(* IEC 61131-3 sources: TSA-FMICS22/ahorn/test/lib_se/file, 7 files *)

(* ---- call_coverage_in_1_cycle_with_change_annotation.st ---- *)
PROGRAM P
VAR_INPUT
    a : INT;
END_VAR
VAR
    f : Fb;
END_VAR
VAR_OUTPUT
    b : BOOL;
END_VAR
    f(x:=a,z=>b);
END_PROGRAM

FUNCTION_BLOCK Fb
VAR_INPUT
    x : INT;
END_VAR
VAR
    y : INT;
END_VAR
VAR_OUTPUT
    z : BOOL;
END_VAR;
    IF x >= 32 THEN
        y := y + change(1, 3);
    ELSE
        y := y;
    END_IF;
    IF y >= 3 THEN
        z := TRUE;
        y := 0;
    ELSE
        z := FALSE;
    END_IF;
END_FUNCTION_BLOCK

(* ---- call_coverage_in_2_cycles.st ---- *)
PROGRAM P
VAR_INPUT
    a : INT;
END_VAR
VAR
    f : Fb;
END_VAR
VAR_OUTPUT
    b : BOOL;
END_VAR
    f(x:=a,z=>b);
END_PROGRAM

FUNCTION_BLOCK Fb
VAR_INPUT
    x : INT;
END_VAR
VAR
    y : INT;
END_VAR
VAR_OUTPUT
    z : BOOL;
END_VAR;
    IF x >= 32 THEN
        y := y + 2;
    ELSE
        y := y;
    END_IF;
    IF y >= 3 THEN
        z := TRUE;
        y := 0;
    ELSE
        z := FALSE;
    END_IF;
END_FUNCTION_BLOCK

(* ---- call_coverage_in_2_cycles_with_change_annotation.st ---- *)
PROGRAM P
VAR_INPUT
    a : INT;
END_VAR
VAR
    f : Fb;
END_VAR
VAR_OUTPUT
    b : BOOL;
END_VAR
    f(x:=a,z=>b);
END_PROGRAM

FUNCTION_BLOCK Fb
VAR_INPUT
    x : INT;
END_VAR
VAR
    y : INT;
END_VAR
VAR_OUTPUT
    z : BOOL;
END_VAR;
    IF x >= 32 THEN
        y := y + change(1, 2);
    ELSE
        y := y;
    END_IF;
    IF y >= 3 THEN
        z := TRUE;
        y := 0;
    ELSE
        z := FALSE;
    END_IF;
END_FUNCTION_BLOCK

(* ---- call_coverage_in_3_cycles.st ---- *)
PROGRAM P
VAR_INPUT
    a : INT;
END_VAR
VAR
    f : Fb;
END_VAR
VAR_OUTPUT
    b : BOOL;
END_VAR
    f(x:=a,z=>b);
END_PROGRAM

FUNCTION_BLOCK Fb
VAR_INPUT
    x : INT;
END_VAR
VAR
    y : INT;
END_VAR
VAR_OUTPUT
    z : BOOL;
END_VAR;
    IF x >= 32 THEN
        y := y + 1;
    ELSE
        y := y;
    END_IF;
    IF y >= 3 THEN
        z := TRUE;
        y := 0;
    ELSE
        z := FALSE;
    END_IF;
END_FUNCTION_BLOCK

(* ---- unreachable_branch_in_call.st ---- *)
PROGRAM P
VAR_INPUT
    a : INT;
END_VAR
VAR
    f : Fb;
END_VAR
VAR_OUTPUT
    b : BOOL;
END_VAR
    f(x:=a,z=>b);
END_PROGRAM

FUNCTION_BLOCK Fb
VAR_INPUT
    x : INT;
END_VAR
VAR
    y : INT;
END_VAR
VAR_OUTPUT
    z : BOOL;
END_VAR;
    IF x >= 32 THEN
        y := y + 1;
    ELSE
        y := y;
    END_IF;
    IF FALSE THEN
        z := TRUE;
        y := 0;
    ELSE
        z := FALSE;
    END_IF;
END_FUNCTION_BLOCK

(* ---- toy_example_kuchta_et_al.st ---- *)
PROGRAM P
VAR_INPUT
    x : INT;
END_VAR
VAR
    y : INT;
    z : INT;
END_VAR
VAR_OUTPUT
    e : BOOL;
    r : INT;
END_VAR
    y := x - 1;
    IF y > 7 THEN
        z := x - 8;
        IF z < 4 THEN
            e := TRUE;
        END_IF;
        r := 0;
    ELSE
        r := 1;
    END_IF;
END_PROGRAM

(* ---- toy_example_kuchta_et_al_with_change_annotation.st ---- *)
PROGRAM P
VAR_INPUT
    x : INT;
END_VAR
VAR
    y : INT;
    z : INT;
END_VAR
VAR_OUTPUT
    e : BOOL;
    r : INT;
END_VAR
    y := change(x - 1, x + 1);
    IF y > 7 THEN
        z := x - 8;
        IF z < 4 THEN
            e := TRUE;
        END_IF;
        r := 0;
    ELSE
        r := 1;
    END_IF;
END_PROGRAM
